// TIA Portal V19 export
DATA_BLOCK "iFB_Press"   // DB20
// stored: InstanceOfName FB_Press, InstanceOfType FB
"FB_Press"
   // VAR_INPUT
   //    Enable : Bool;
   //    Power : Bool;
   //    Emg : Bool;
   //    Ready : Bool;
   //    MainMotor : Bool;
   //    Start_Cycle : Bool;
   //    Stop_Motor : Bool;
   //    SensorTop : Bool;
   // END_VAR
   // VAR_OUTPUT
   //    Busy : Bool;
   //    Done : Bool;
   //    Error : Bool;
   //    Cycle : Bool;
   //    Switch_Off : Bool;
   //    Switch_SafetyStroke : Bool;
   //    Motor_Start : Bool;
   //    Motor_Stop : Bool;
   //    Power_On : Bool;
   //    Power_Off : Bool;
   //    Reset : Bool;
   // END_VAR
   // VAR
   //    iStage : Int;
   //    iCycle : Int;
   //    PressReady : Bool;
   // END_VAR
BEGIN
END_DATA_BLOCK
